(* IEC 61131-3 sources: llm-plc-st-eval/data/definitivo/qwen2.5-coder_14b/A6/zero_shot, 3 files *)

(* ---- ejec_1.st ---- *)
```structured-text
FUNCTION_BLOCK FB_Modos
VAR_INPUT
    selector : INT;          // Selector de modo (0: automático, 1: manual, 2: mantenimiento)
    estadoSeguro : BOOL;      // Estado de seguridad activo/inactivo
    cmdAuto : ARRAY[0..7] OF BOOL; // Comandos automáticos para los actuadores
    cmdManual : ARRAY[0..7] OF BOOL; // Comandos manuales para los actuadores
    idxForzado : INT;        // Índice del actuador a forzar
    valorForzado : BOOL;     // Valor a forzar en el actuador
    confirmarForzado : BOOL; // Confirmación de forzado
END_VAR

VAR_OUTPUT
    modoActivo : INT;        // Modo activo (0: automático, 1: manual, 2: mantenimiento)
    actuador : ARRAY[0..7] OF BOOL; // Estado de los actuadores
END_VAR

VAR
    modoVigente : INT := 1;  // Modo vigente inicializado a manual (1)
    forzado : ARRAY[0..7] OF BOOL; // Estado de forzado de los actuadores
END_VAR

METHOD Update : VOID
VAR
    i : INT;
END_VAR

    // Mantener el modo vigente si el selector está fuera de rango
    IF selector < 0 OR selector > 2 THEN
        modoActivo := modoVigente;
    ELSE
        modoActivo := selector;
    END_IF;

    // Cambiar el modo vigente solo si estadoSeguro está activo
    IF estadoSeguro THEN
        modoVigente := modoActivo;
    END_IF;

    // Manejo de los actuadores según el modo activo
    CASE modoActivo OF
        0: // Modo automático
            FOR i := 0 TO 7 DO
                actuador[i] := cmdAuto[i];
            END_FOR;
        1: // Modo manual
            FOR i := 0 TO 7 DO
                actuador[i] := cmdManual[i];
            END_FOR;
        2: // Modo mantenimiento
            FOR i := 0 TO 7 DO
                actuador[i] := FALSE;
            END_FOR;
            IF confirmarForzado THEN
                IF idxForzado >= 0 AND idxForzado <= 7 THEN
                    actuador[idxForzado] := valorForzado;
                    forzado[idxForzado] := TRUE;
                END_IF;
            END_IF;
            IF NOT estadoSeguro THEN
                FOR i := 0 TO 7 DO
                    forzado[i] := FALSE;
                END_FOR;
            END_IF;
    END_CASE;

    // Anular forzados al salir del modo mantenimiento
    IF modoActivo <> 2 THEN
        FOR i := 0 TO 7 DO
            forzado[i] := FALSE;
        END_FOR;
    END_IF;
END_METHOD

// Llamada al método Update en cada ciclo
Update();
END_FUNCTION_BLOCK
```

(* ---- ejec_2.st ---- *)
```iec
FUNCTION_BLOCK FB_Modos
VAR_INPUT
    selector : INT;          // Selector de modo (0: Automático, 1: Manual, 2: Mantenimiento)
    estadoSeguro : BOOL;      // Estado de seguridad activo/inactivo
    cmdAuto : ARRAY[0..7] OF BOOL; // Comandos automáticos para los actuadores
    cmdManual : ARRAY[0..7] OF BOOL; // Comandos manuales para los actuadores
    idxForzado : INT;        // Índice del actuador a forzar (0-7)
    valorForzado : BOOL;     // Valor a forzar en el actuador
    confirmarForzado : BOOL; // Confirmación de forzado
END_VAR

VAR_OUTPUT
    modoActivo : INT;         // Modo activo (0: Automático, 1: Manual, 2: Mantenimiento)
    actuador : ARRAY[0..7] OF BOOL; // Estado de los actuadores
END_VAR

VAR
    modoVigente : INT := 1;  // Modo vigente inicializado a Manual (1)
    forzado : ARRAY[0..7] OF BOOL; // Estado de forzado de los actuadores
    forzadoActivo : BOOL := FALSE; // Indica si hay algún forzado activo
END_VAR

METHOD Update : VOID
VAR
    i : INT;
END_VAR

    // Mantener el modo vigente si el selector está fuera de rango
    IF selector < 0 OR selector > 2 THEN
        modoActivo := modoVigente;
    ELSE
        modoActivo := selector;
    END_IF;

    // Cambiar el modo vigente solo si estadoSeguro está activo
    IF estadoSeguro THEN
        modoVigente := modoActivo;
    END_IF;

    // Actualizar los actuadores según el modo activo
    CASE modoActivo OF
        0: // Modo Automático
            FOR i := 0 TO 7 DO
                actuador[i] := cmdAuto[i];
            END_FOR;
        1: // Modo Manual
            FOR i := 0 TO 7 DO
                actuador[i] := cmdManual[i];
            END_FOR;
        2: // Modo Mantenimiento
            FOR i := 0 TO 7 DO
                actuador[i] := FALSE;
            END_FOR;
            IF confirmarForzado THEN
                IF idxForzado >= 0 AND idxForzado <= 7 THEN
                    actuador[idxForzado] := valorForzado;
                    forzado[idxForzado] := TRUE;
                    forzadoActivo := TRUE;
                END_IF;
            END_IF;
    END_CASE;

    // Anular los forzados si estadoSeguro se desactiva o se sale del modo mantenimiento
    IF NOT estadoSeguro OR modoActivo <> 2 THEN
        FOR i := 0 TO 7 DO
            forzado[i] := FALSE;
            actuador[i] := FALSE;
        END_FOR;
        forzadoActivo := FALSE;
    END_IF;

END_METHOD

END_FUNCTION_BLOCK
```

(* ---- ejec_3.st ---- *)
```pascal
FUNCTION_BLOCK FB_Modos
VAR_INPUT
    selector : INT;          // Selector de modo (0: automático, 1: manual, 2: mantenimiento)
    estadoSeguro : BOOL;      // Estado de seguridad activo/inactivo
    cmdAuto : ARRAY[0..7] OF BOOL;  // Comandos para modo automático
    cmdManual : ARRAY[0..7] OF BOOL;  // Comandos para modo manual
    idxForzado : INT;        // Índice del actuador a forzar en modo mantenimiento
    valorForzado : BOOL;      // Valor a forzar en el actuador seleccionado
    confirmarForzado : BOOL;  // Confirmación de forzado
END_VAR

VAR_OUTPUT
    modoActivo : INT;         // Modo de operación activo
    actuador : ARRAY[0..7] OF BOOL;  // Estado de los actuadores
END_VAR

VAR
    modoAnterior : INT;       // Modo anterior para comparación
    forzado : ARRAY[0..7] OF BOOL;  // Estado de forzado de los actuadores
END_VAR

// Inicialización en el arranque
IF NOT estadoSeguro THEN
    modoActivo := 1;  // Modo manual por defecto
ELSE
    modoAnterior := modoActivo;
    CASE selector OF
        0..2: modoActivo := selector;  // Cambio de modo si el selector está en un valor válido
        ELSE modoActivo := modoAnterior;  // Mantener modo anterior si el selector está fuera de rango
    END_CASE;
END_IF;

// Gestión de los actuadores según el modo
CASE modoActivo OF
    0:  // Modo automático
        FOR i := 0 TO 7 DO
            actuador[i] := cmdAuto[i];
        END_FOR;
    1:  // Modo manual
        FOR i := 0 TO 7 DO
            actuador[i] := cmdManual[i];
        END_FOR;
    2:  // Modo mantenimiento
        IF NOT estadoSeguro THEN
            FOR i := 0 TO 7 DO
                actuador[i] := FALSE;
                forzado[i] := FALSE;
            END_FOR;
        ELSE
            IF confirmarForzado THEN
                IF idxForzado >= 0 AND idxForzado <= 7 THEN
                    actuador[idxForzado] := valorForzado;
                    forzado[idxForzado] := TRUE;
                END_IF;
            END_IF;
        END_IF;
END_CASE;

// Anulación de forzados al salir del modo mantenimiento
IF modoAnterior = 2 AND modoActivo <> 2 THEN
    FOR i := 0 TO 7 DO
        forzado[i] := FALSE;
    END_FOR;
END_IF;

// Anulación de forzados si estadoSeguro se desactiva durante el mantenimiento
IF modoActivo = 2 AND NOT estadoSeguro THEN
    FOR i := 0 TO 7 DO
        actuador[i] := FALSE;
        forzado[i] := FALSE;
    END_FOR;
END_IF;

modoAnterior := modoActivo;
END_FUNCTION_BLOCK
```
